FUNCTION_BLOCK FB_Scale
VAR_INPUT
    RawValue : INT;       
    RawMin   : REAL := 0.0;     
    RawMax   : REAL := 32767.0; 
    PhysMin  : REAL;      
    PhysMax  : REAL;      
END_VAR

VAR_OUTPUT
    ScaledValue : REAL;   
END_VAR

// Error handling to prevent division by zero.
IF (RawMax - RawMin) <> 0.0 THEN
    ScaledValue :=  PhysMin + (PhysMax - PhysMin) * (INT_TO_REAL(RawValue) - RawMin) / (RawMax - RawMin);
ELSE
    ScaledValue := PhysMin;
END_IF

END_FUNCTION_BLOCK

(* stored: Version 1.1.0.1, ProductVersion 3.1.4026.21
   POU FB_Scale: Id {da1442ee-1458-4201-b087-62b994f875f2}, SpecialFunc None *)
